// TIA Portal V20 export
// export: Created 2026-10-20T18:54:30.6966194Z, ExportSetting None, DisplayName Totally Integrated Automation Portal, DisplayVersion V20 Update 6, DisplayName TIA Portal Openness, DisplayVersion V20 Update 6, DisplayName TIA Portal Version Control Interface, DisplayVersion V20 Update 6, DisplayName SINAMICS Startdrive Advanced, DisplayVersion V20 SP1, DisplayName SINAMICS Startdrive G130, G150, S120, S150, SINAMICS MV, G220, S200, S210, DisplayVersion V20 SP1, DisplayName SINAMICS Startdrive G110M, G120, G120C, G120D, G120P, G115D, DisplayVersion V20 SP1, DisplayName STEP 7 Professional, DisplayVersion V20 Update 6, DisplayName STEP 7 Safety, DisplayVersion V20 Update 2, DisplayName WinCC Basic/Comfort/Advanced, DisplayVersion V20 Update 6, DisplayName WinCC Unified, DisplayVersion V20 Update 6
VAR_GLOBAL   // PLC tag table "VTD_HMI_IO"
   VTD_DP1_Retracted_HMI AT %M8.2 : Bool;
   VTD_DP2_Extended_HMI AT %M8.1 : Bool;
   VTD_Upper_Overtravel_HMI AT %M19.3 : Bool;
   VTD_DP1_Extended_HMI AT %M6.2 : Bool;
   VTD_DP2_Retracted_HMI AT %M8.3 : Bool;
   VTD_Lower_Overtravel_HMI AT %M19.2 : Bool;
   VTD_Level_Detect1_HMI AT %M4.7 : Bool;
   VTD_Lower_Limit_HMI AT %M4.6 : Bool;
   VTD_Ultimate_Creep_HMI AT %M5.2 : Bool;
   VTD_Upper_Limet_HMI AT %M3.1 : Bool;
   VTD_Level_Detect2_HMI AT %M5.0 : Bool;
   VTD_Ultimate_Slow_HMI AT %M5.1 : Bool;
   VTD_Upper_Limet_Bypass_HMI AT %M60.4 : Bool;
   VTD_Lower_Limit_Bypass_HMI AT %M60.5 : Bool;
   VTD_Upper_Overtravel_Bypass_HMI AT %M60.6 : Bool;
   VTD_Lower_Overtravel_Bypass_HMI AT %M60.7 : Bool;
   Chain_Slack_1_Bypass_HMI AT %M61.0 : Bool;
   Chain_Slack_2_Bypass_HMI AT %M61.1 : Bool;
   Chain_Slack_3_Bypass_HMI AT %M61.2 : Bool;
   Chain_Slack_4_Bypass_HMI AT %M61.3 : Bool;
END_VAR
